(* IEC 61131-3 sources: lab-assay-lims/projects/plc-control-panel-design/design, 1 file *)

(* ---- source-line.st ---- *)
(* Generated by OpenPLC editor 6a8e930a914e4421e8fa05966b31eb371b439243; source: plc/line.xml. *)
PROGRAM FillingLine
  VAR_INPUT
    Start : BOOL;
    Stop : BOOL;
    Reset : BOOL;
    EStopOK : BOOL;
    GuardClosed : BOOL;
    TankOK : BOOL;
    BottleAtFill : BOOL;
    ExitSensor : BOOL;
    JamSwitch : BOOL;
  END_VAR
  VAR_OUTPUT
    Run : BOOL;
    Conveyor : BOOL;
    Valve : BOOL;
    Alarm : BOOL;
    BatchDone : BOOL;
    FillBlocked : BOOL;
  END_VAR
  VAR
    Fault : BOOL;
    Filled : BOOL;
    StartEdge : R_TRIG;
    ExitEdge : R_TRIG;
    BatchCount : CTU;
    JamTimer : TON;
    FillTimer : TON;
    FillClearTimer : TON;
  END_VAR

  StartEdge(CLK := Start);
  ExitEdge(CLK := ExitSensor);
  BatchCount(CU := Run AND ExitEdge.Q, R := Reset, PV := 5);
  JamTimer(IN := NOT(ExitSensor) AND Conveyor, PT := T#3000ms);
  FillClearTimer(IN := BottleAtFill AND Filled AND Run, PT := T#1000ms);
  FillTimer(IN := NOT(Filled) AND BottleAtFill AND Run, PT := T#1000ms);
  FillBlocked := FillClearTimer.Q OR (BottleAtFill OR NOT(Reset)) AND FillBlocked;
  Fault := FillBlocked OR JamSwitch OR JamTimer.Q OR NOT(EStopOK) OR NOT(GuardClosed) OR NOT(TankOK) OR (BottleAtFill OR NOT(Reset)) AND Fault OR NOT(Filled) AND BottleAtFill AND Run AND Stop;
  Run := NOT(BatchCount.Q) AND NOT(Fault) AND TankOK AND GuardClosed AND EStopOK AND NOT(Stop) AND (Run OR StartEdge.Q);
  Filled := Run AND BottleAtFill AND (FillTimer.Q OR Filled);
  Conveyor := (Filled OR NOT(BottleAtFill)) AND Run;
  Valve := NOT(Filled) AND BottleAtFill AND Run;
  Alarm := Fault;
  BatchDone := BatchCount.Q;
END_PROGRAM

CONFIGURATION LineConfig

  RESOURCE CPU ON PLC
    TASK Scan(INTERVAL := T#50ms,PRIORITY := 0);
    PROGRAM Line WITH Scan : FillingLine;
  END_RESOURCE
END_CONFIGURATION
